(* IEC 61131-3 sources: sis-interlock-demo/pytests/golden/mini/src/DUTs/Generated, 1 file *)

(* ---- ST_SisIo.dut.st ---- *)
// AUTO-GENERATED by cemgen 1.0.0 — не редактировать: правьте матрицу и запустите
//   python -m cemgen generate <файл матрицы .csv или .xlsx>
// Матрица: TEST-U301-CEM, объект U-301, ревизия 1 от 2026-10-16, SHA-256 сетки 9067fda96ae55e67
// Назначение: образ ввода-вывода ПАЗ объекта U-301: токи датчиков 4–20 мА, дискретные входы с
//             контролем линии, ключи и кнопка, выходы-разрешения xQ* (TRUE — под напряжением).
//             Поля — по тегам матрицы (DESIGN.md, 9.3), порядок — первое появление каналов, затем
//             ключи и выходы.
// Автор:      pytest; код — генератор cemgen
// Версия:     1.0.0
// Документ:   docs/DESIGN.md, раздел «10. Генератор cemgen»; docs/cause_effect_matrix.md
// ВНИМАНИЕ:   код демонстрационный и не предназначен для систем безопасности. Реальная ПАЗ требует
//             определения SIL, сертифицированных аппаратных и программных средств и валидации по
//             ГОСТ Р МЭК 61511.
{attribute 'qualified_only'}
TYPE ST_SisIo :
STRUCT
    // --- 1 TSH301: Температура высокая (ai, 1oo1) ---
    rTT301_mA  : REAL;   // TT301, мА: шкала 0…100 °C; 1 TSH301
    // --- 2 PSL302: Давление низкое (di, 2oo2) ---
    xPS302A    : BOOL;   // PS302A: норма 1; 2 PSL302
    xPS302A_Ok : BOOL;   // PS302A: контроль линии, TRUE — исправна
    xPS302B    : BOOL;   // PS302B: норма 1; 2 PSL302
    xPS302B_Ok : BOOL;   // PS302B: контроль линии, TRUE — исправна
    // --- 3 XS303: Внешний останов (ext, —) ---
    xXS303     : BOOL;   // XS303: внешнее требование, норма 0; 3 XS303
    // --- выходы ПАЗ: разрешения, обесточивание на срабатывание ---
    xQXV301    : BOOL;   // XV301: разрешение, TRUE — под напряжением; FALSE — закрыт
    xQM302     : BOOL;   // M302: разрешение, TRUE — под напряжением; FALSE — остановлен
END_STRUCT
END_TYPE
